(* IEC 61131-3 sources: llm-plc-st-eval/codesys/dobles/B8, 9 files *)

(* ---- 01_Correcta.st ---- *)
(* DOBLE DE PRUEBA B8/Correcta - NO ES CORPUS. Esperado: veredicto 1 *)
FUNCTION_BLOCK FB_Puerta
VAR_INPUT
    puertaAbierta : BOOL;
    reset : BOOL;
END_VAR
VAR_OUTPUT
    aviso : BOOL;
    nAperturas : INT;
END_VAR
VAR
    prev : BOOL;
END_VAR
IF reset THEN
    nAperturas := 0;
ELSIF puertaAbierta AND NOT prev THEN
    nAperturas := nAperturas + 1;
END_IF
prev := puertaAbierta;
aviso := nAperturas >= 5;
END_FUNCTION_BLOCK

(* ---- 02_CuentaPorNivel.st ---- *)
(* DOBLE DE PRUEBA B8/CuentaPorNivel - NO ES CORPUS. Esperado: veredicto 2, falla en el paso 1 *)
FUNCTION_BLOCK FB_Puerta
VAR_INPUT
    puertaAbierta : BOOL;
    reset : BOOL;
END_VAR
VAR_OUTPUT
    aviso : BOOL;
    nAperturas : INT;
END_VAR
VAR
    prev : BOOL;
END_VAR
IF reset THEN
    nAperturas := 0;
ELSIF puertaAbierta THEN
    nAperturas := nAperturas + 1;
END_IF
prev := puertaAbierta;
aviso := nAperturas >= 5;
END_FUNCTION_BLOCK

(* ---- 03_CuentaFlancoBajada.st ---- *)
(* DOBLE DE PRUEBA B8/CuentaFlancoBajada - NO ES CORPUS. Esperado: veredicto 2, falla en el paso 1 *)
FUNCTION_BLOCK FB_Puerta
VAR_INPUT
    puertaAbierta : BOOL;
    reset : BOOL;
END_VAR
VAR_OUTPUT
    aviso : BOOL;
    nAperturas : INT;
END_VAR
VAR
    prev : BOOL;
END_VAR
IF reset THEN
    nAperturas := 0;
ELSIF prev AND NOT puertaAbierta THEN
    nAperturas := nAperturas + 1;
END_IF
prev := puertaAbierta;
aviso := nAperturas >= 5;
END_FUNCTION_BLOCK

(* ---- 04_UmbralCuatro.st ---- *)
(* DOBLE DE PRUEBA B8/UmbralCuatro - NO ES CORPUS. Esperado: veredicto 2, falla en el paso 4 *)
FUNCTION_BLOCK FB_Puerta
VAR_INPUT
    puertaAbierta : BOOL;
    reset : BOOL;
END_VAR
VAR_OUTPUT
    aviso : BOOL;
    nAperturas : INT;
END_VAR
VAR
    prev : BOOL;
END_VAR
IF reset THEN
    nAperturas := 0;
ELSIF puertaAbierta AND NOT prev THEN
    nAperturas := nAperturas + 1;
END_IF
prev := puertaAbierta;
aviso := nAperturas >= 4;
END_FUNCTION_BLOCK

(* ---- 05_UmbralSeis.st ---- *)
(* DOBLE DE PRUEBA B8/UmbralSeis - NO ES CORPUS. Esperado: veredicto 2, falla en el paso 5 *)
FUNCTION_BLOCK FB_Puerta
VAR_INPUT
    puertaAbierta : BOOL;
    reset : BOOL;
END_VAR
VAR_OUTPUT
    aviso : BOOL;
    nAperturas : INT;
END_VAR
VAR
    prev : BOOL;
END_VAR
IF reset THEN
    nAperturas := 0;
ELSIF puertaAbierta AND NOT prev THEN
    nAperturas := nAperturas + 1;
END_IF
prev := puertaAbierta;
aviso := nAperturas > 5;
END_FUNCTION_BLOCK

(* ---- 06_AvisoSoloEnCinco.st ---- *)
(* DOBLE DE PRUEBA B8/AvisoSoloEnCinco - NO ES CORPUS. Esperado: veredicto 2, falla en el paso 6 *)
FUNCTION_BLOCK FB_Puerta
VAR_INPUT
    puertaAbierta : BOOL;
    reset : BOOL;
END_VAR
VAR_OUTPUT
    aviso : BOOL;
    nAperturas : INT;
END_VAR
VAR
    prev : BOOL;
END_VAR
IF reset THEN
    nAperturas := 0;
ELSIF puertaAbierta AND NOT prev THEN
    nAperturas := nAperturas + 1;
END_IF
prev := puertaAbierta;
aviso := nAperturas = 5;
END_FUNCTION_BLOCK

(* ---- 07_SaturaEnCinco.st ---- *)
(* DOBLE DE PRUEBA B8/SaturaEnCinco - NO ES CORPUS. Esperado: veredicto 2, falla en el paso 6 *)
FUNCTION_BLOCK FB_Puerta
VAR_INPUT
    puertaAbierta : BOOL;
    reset : BOOL;
END_VAR
VAR_OUTPUT
    aviso : BOOL;
    nAperturas : INT;
END_VAR
VAR
    prev : BOOL;
END_VAR
IF reset THEN
    nAperturas := 0;
ELSIF puertaAbierta AND NOT prev AND nAperturas < 5 THEN
    nAperturas := nAperturas + 1;
END_IF
prev := puertaAbierta;
aviso := nAperturas >= 5;
END_FUNCTION_BLOCK

(* ---- 08_ResetNoApagaAviso.st ---- *)
(* DOBLE DE PRUEBA B8/ResetNoApagaAviso - NO ES CORPUS. Esperado: veredicto 2, falla en el paso 7 *)
FUNCTION_BLOCK FB_Puerta
VAR_INPUT
    puertaAbierta : BOOL;
    reset : BOOL;
END_VAR
VAR_OUTPUT
    aviso : BOOL;
    nAperturas : INT;
END_VAR
VAR
    prev : BOOL;
END_VAR
IF reset THEN
    nAperturas := 0;
ELSIF puertaAbierta AND NOT prev THEN
    nAperturas := nAperturas + 1;
END_IF
prev := puertaAbierta;
aviso := aviso OR nAperturas >= 5;
END_FUNCTION_BLOCK

(* ---- 09_ResetSoloAviso.st ---- *)
(* DOBLE DE PRUEBA B8/ResetSoloAviso - NO ES CORPUS. Esperado: veredicto 2, falla en el paso 7 *)
FUNCTION_BLOCK FB_Puerta
VAR_INPUT
    puertaAbierta : BOOL;
    reset : BOOL;
END_VAR
VAR_OUTPUT
    aviso : BOOL;
    nAperturas : INT;
END_VAR
VAR
    prev : BOOL;
END_VAR
IF reset THEN
    aviso := FALSE;
ELSIF puertaAbierta AND NOT prev THEN
    nAperturas := nAperturas + 1;
END_IF
prev := puertaAbierta;
IF NOT reset THEN
    aviso := nAperturas >= 5;
END_IF
END_FUNCTION_BLOCK
